(* IEC 61131-3 sources: llm-plc-st-eval/data/definitivo/gpt-4o-2024-08-06/B4/zero_shot, 3 files *)

(* ---- ejec_1.st ---- *)
```pascal
FUNCTION_BLOCK FB_Giro
VAR_INPUT
    btnFwd : BOOL;   // Botón para giro en sentido horario
    btnRev : BOOL;   // Botón para giro en sentido antihorario
    btnParo : BOOL;  // Botón de paro
END_VAR

VAR_OUTPUT
    fwd : BOOL;      // Salida para giro en sentido horario
    rev : BOOL;      // Salida para giro en sentido antihorario
END_VAR

VAR
    estado : INT;    // Estado del motor: 0 = Paro, 1 = Horario, 2 = Antihorario
END_VAR

// Inicialización de salidas
fwd := FALSE;
rev := FALSE;

// Lógica de control del motor
IF btnParo THEN
    estado := 0; // Cambiar a estado de paro
ELSIF btnFwd AND (estado = 0) THEN
    estado := 1; // Cambiar a estado de giro horario
ELSIF btnRev AND (estado = 0) THEN
    estado := 2; // Cambiar a estado de giro antihorario
END_IF

// Actualización de salidas según el estado
CASE estado OF
    0: // Paro
        fwd := FALSE;
        rev := FALSE;
    1: // Giro horario
        fwd := TRUE;
        rev := FALSE;
    2: // Giro antihorario
        fwd := FALSE;
        rev := TRUE;
END_CASE
END_FUNCTION_BLOCK
```

Este código implementa la lógica de inversión de giro de un motor, asegurando que las salidas `fwd` y `rev` nunca estén activas al mismo tiempo y que el motor pase por el estado de paro antes de cambiar de dirección.

(* ---- ejec_2.st ---- *)
```pascal
FUNCTION_BLOCK FB_Giro
VAR_INPUT
    btnFwd : BOOL;   // Botón para giro en sentido horario
    btnRev : BOOL;   // Botón para giro en sentido antihorario
    btnParo : BOOL;  // Botón para detener el motor
END_VAR

VAR_OUTPUT
    fwd : BOOL;      // Salida para giro en sentido horario
    rev : BOOL;      // Salida para giro en sentido antihorario
END_VAR

VAR
    estado : INT;    // Estado actual del motor: 0 = Paro, 1 = Fwd, 2 = Rev
END_VAR

// Inicialización del estado
estado := 0;

// Lógica de control del motor
IF btnParo THEN
    // Si se presiona el botón de paro, detener el motor
    estado := 0;
ELSIF btnFwd AND (estado = 0) THEN
    // Si se presiona el botón de avance y el motor está parado, girar en sentido horario
    estado := 1;
ELSIF btnRev AND (estado = 0) THEN
    // Si se presiona el botón de retroceso y el motor está parado, girar en sentido antihorario
    estado := 2;
END_IF

// Actualización de las salidas según el estado
CASE estado OF
    0: // Estado de paro
        fwd := FALSE;
        rev := FALSE;
    1: // Estado de giro en sentido horario
        fwd := TRUE;
        rev := FALSE;
    2: // Estado de giro en sentido antihorario
        fwd := FALSE;
        rev := TRUE;
END_CASE

END_FUNCTION_BLOCK
```

Este código implementa la lógica de inversión de giro de un motor, asegurando que el motor pase por un estado de paro antes de cambiar de dirección. Las salidas `fwd` y `rev` nunca estarán activas al mismo tiempo, cumpliendo con los requisitos especificados.

(* ---- ejec_3.st ---- *)
```pascal
FUNCTION_BLOCK FB_Giro
VAR_INPUT
    btnFwd : BOOL;   // Botón para giro en sentido horario
    btnRev : BOOL;   // Botón para giro en sentido antihorario
    btnParo : BOOL;  // Botón de paro
END_VAR

VAR_OUTPUT
    fwd : BOOL;      // Salida para giro en sentido horario
    rev : BOOL;      // Salida para giro en sentido antihorario
END_VAR

VAR
    estado : INT;    // Estado del motor: 0 = Parado, 1 = Horario, 2 = Antihorario
END_VAR

// Inicialización de salidas
fwd := FALSE;
rev := FALSE;

// Lógica de control
IF btnParo THEN
    // Si se presiona el botón de paro, el motor se detiene
    estado := 0;
ELSIF btnFwd AND (estado = 0) THEN
    // Si se presiona el botón de giro horario y el motor está parado
    estado := 1;
ELSIF btnRev AND (estado = 0) THEN
    // Si se presiona el botón de giro antihorario y el motor está parado
    estado := 2;
END_IF

// Actualización de salidas según el estado
CASE estado OF
    0: // Parado
        fwd := FALSE;
        rev := FALSE;
    1: // Giro horario
        fwd := TRUE;
        rev := FALSE;
    2: // Giro antihorario
        fwd := FALSE;
        rev := TRUE;
END_CASE;

END_FUNCTION_BLOCK
```

Este código implementa la lógica para controlar la inversión de giro de un motor, asegurando que nunca se activen ambas salidas simultáneamente y que siempre se pase por el estado de paro antes de cambiar de dirección.
